(* IEC 61131-3 sources: moqui-plc/rust-plc/interfaces/codesys-iiot, 3 files *)

(* ---- json.st ---- *)
(* CODESYS IIoT JSON API used by moqui-plc (library namespace JSON).
 *
 * Interface declarations only (no implementation), for type checking with a
 * non-CODESYS compiler. The vendor library is object oriented (methods on
 * function blocks); the declarations mirror only the calls moqui-plc makes.
 *)

TYPE JSON_ERROR : (NO_ERROR, INVALID_INPUT, NO_MEMORY, NOT_FOUND, PARSE_ERROR); END_TYPE
TYPE JSONType : (JSON_OBJECT, JSON_ARRAY, KEY, VALUE); END_TYPE

TYPE JSONValue :
STRUCT
    wsValue : WSTRING(255);
    lrValue : LREAL;
    diValue : DINT;
    xValue : BOOL;
END_STRUCT
END_TYPE

TYPE JSONElement :
STRUCT
    eType : JSONType;
    diIndex : DINT;
    diParentIndex : DINT;
    value : JSONValue;
END_STRUCT
END_TYPE

FUNCTION_BLOCK JSONData
METHOD Clear
END_METHOD
METHOD GetElementByIndex : JSON_ERROR
VAR_INPUT
    diIndex : DINT;
END_VAR
VAR_OUTPUT
    jsonElement : JSONElement;
END_VAR
END_METHOD
METHOD GetChildren : JSON_ERROR
VAR_INPUT
    diIndex : DINT;
    pResult : POINTER TO JSONElement;
    udiMaxSize : UDINT;
END_VAR
VAR_OUTPUT
    udiResultSize : UDINT;
END_VAR
END_METHOD
END_FUNCTION_BLOCK

FUNCTION_BLOCK JSONDataFactory
METHOD Create : POINTER TO JSONData
VAR_OUTPUT
    eError : JSON_ERROR;
END_VAR
END_METHOD
END_FUNCTION_BLOCK

FUNCTION_BLOCK JSONBuilder
VAR_INPUT
    pJsonData : POINTER TO JSONData;
END_VAR
VAR_OUTPUT
    diRootObj : DINT;
END_VAR
METHOD Reset
END_METHOD
METHOD SetKeyWithObject : DINT
VAR_INPUT
    wsKey : WSTRING;
    diParentIndex : DINT;
END_VAR
END_METHOD
METHOD SetKeyWithValue : DINT
VAR_INPUT
    wsKey : WSTRING;
    value : ANY;
    diParentIndex : DINT;
END_VAR
END_METHOD
END_FUNCTION_BLOCK

FUNCTION_BLOCK JSONByteArrayWriter
VAR_INPUT
    xExecute : BOOL;
    xAsyncMode : BOOL;
    pwData : POINTER TO WORD;
    udiSize : UDINT;
    wsLineBreak : WSTRING(2);
END_VAR
VAR_IN_OUT
    jsonData : JSONData;
END_VAR
VAR_OUTPUT
    xDone : BOOL;
    xBusy : BOOL;
    xError : BOOL;
    eError : JSON_ERROR;
END_VAR
END_FUNCTION_BLOCK

FUNCTION_BLOCK JSONByteArrayReader
VAR_INPUT
    xExecute : BOOL;
    xAsyncMode : BOOL;
    pwData : POINTER TO WORD;
END_VAR
VAR_IN_OUT
    jsonData : JSONData;
END_VAR
VAR_OUTPUT
    xDone : BOOL;
    xBusy : BOOL;
    xError : BOOL;
    eError : JSON_ERROR;
END_VAR
END_FUNCTION_BLOCK

(* ---- mqtt.st ---- *)
(* CODESYS IIoT MQTT client API used by moqui-plc (library namespace MQTT).
 *
 * Interface declarations only (no implementation), for type checking with a
 * non-CODESYS compiler. Only the members moqui-plc uses are declared. A Rust
 * runtime would implement them on top of an MQTT 5 client crate.
 *)

TYPE MQTT_VERSION : (V3_1_1 := 4, V5 := 5); END_TYPE
TYPE MQTT_QOS : (QoS0, QoS1, QoS2); END_TYPE
TYPE MQTT_RETAIN_HANDLING : (On_Subscribe, If_Not_Exists, Not_Exists); END_TYPE
TYPE COMMUNICATION_MODE : (TCP, WEBSOCKET); END_TYPE
TYPE FILTER_MODE : (FILTER_OFF, FILTER_ON); END_TYPE
TYPE MQTT_ERROR : (NO_ERROR, TIMEOUT, CONNECTION_REFUSED, DISCONNECTED, PROTOCOL_ERROR); END_TYPE

(* Library parameters (CODESYS: MQTT.MQTTParam). Values are runtime specific. *)
VAR_GLOBAL CONSTANT
    g_udiMaxPacketSize : UDINT := 268435455;
    g_udiMaxUserProperties : UDINT := 8;
END_VAR

TYPE MQTTConnectProperties :
STRUCT
    udiSessionExpiryInterval : UDINT;
    udiMaximumPacketSize : UDINT;
END_STRUCT
END_TYPE

TYPE MQTTWillProperties :
STRUCT
    bPayloadFormatIndicator : BYTE;
    udiMessageExpiryInterval : UDINT;
    wsContentType : WSTRING;
    udiWillDelayInterval : UDINT;
END_STRUCT
END_TYPE

TYPE MQTTPublishProperties :
STRUCT
    bPayloadFormatIndicator : BYTE;
    udiMessageExpiryInterval : UDINT;
    wsContentType : WSTRING;
END_STRUCT
END_TYPE

TYPE MQTTSubscribeProperties :
STRUCT
    udiSubscriptionIdentifier : UDINT;
    xNoLocalOption : BOOL;
    xRetainAsPublished : BOOL;
    eRetainHandling : MQTT_RETAIN_HANDLING;
END_STRUCT
END_TYPE

FUNCTION_BLOCK MQTTClient
VAR_INPUT
    xEnable : BOOL;
    sHostname : STRING(255);
    uiPort : UINT;
    eCommunicationMode : COMMUNICATION_MODE;
    sWebSocketUrl : STRING(255);
    itfTLSContext : ITLSContext;
    eMQTTVersion : MQTT_VERSION;
    sClientId : STRING(255);
    wsUsername : WSTRING(255);
    wsPassword : WSTRING(255);
    uiKeepAlive : UINT;
    xCleanSession : BOOL;
    udiTimeOut : UDINT;
    tPingInterval : TIME;
    wsWillTopic : WSTRING(1024);
    pbWillMessage : POINTER TO BYTE;
    uiWillMessageSize : UINT;
    eWillQoS : MQTT_QOS;
    xWillRetain : BOOL;
    mQTTConnectProperties : MQTTConnectProperties;
    mQTTWillProperties : MQTTWillProperties;
END_VAR
VAR_OUTPUT
    xConnectedToBroker : BOOL;
    xBusy : BOOL;
    xError : BOOL;
    eMQTTError : MQTT_ERROR;
END_VAR
END_FUNCTION_BLOCK

FUNCTION_BLOCK MQTTPublish
VAR_INPUT
    xExecute : BOOL;
    mqttClient : REF_TO MQTTClient;
    wsTopicName : WSTRING(1024);
    pbPayload : POINTER TO BYTE;
    udiPayloadSize : UDINT;
    eQoS : MQTT_QOS;
    xRetain : BOOL;
    xReDelivery : BOOL;
    udiTimeOut : UDINT;
    mQTTPublishProperties : MQTTPublishProperties;
END_VAR
VAR_OUTPUT
    xDone : BOOL;
    xBusy : BOOL;
    xError : BOOL;
    eMQTTError : MQTT_ERROR;
END_VAR
END_FUNCTION_BLOCK

FUNCTION_BLOCK MQTTSubscribe
VAR_INPUT
    xEnable : BOOL;
    mqttClient : REF_TO MQTTClient;
    wsTopicFilter : WSTRING(1024);
    eFilterMode : FILTER_MODE;
    eSubscribeQoS : MQTT_QOS;
    pbPayload : POINTER TO BYTE;
    udiMaxPayloadSize : UDINT;
    udiTimeout : UDINT;
    mQTTSubscribeProperties : MQTTSubscribeProperties;
END_VAR
VAR_OUTPUT
    xDone : BOOL;
    xBusy : BOOL;
    xError : BOOL;
    eMQTTError : MQTT_ERROR;
    xSubscribeActive : BOOL;
    xReceived : BOOL;
    wsLastTopic : WSTRING(1024);
END_VAR
END_FUNCTION_BLOCK

(* ---- tls.st ---- *)
(* CODESYS Net Base Services TLS types used by moqui-plc (library namespace NBS).
 *
 * Interface declarations only (no implementation), for type checking with a
 * non-CODESYS compiler.
 *)

TYPE PURPOSE : (CLIENT_SIDE, SERVER_SIDE); END_TYPE

TYPE CIPHER_LIST :
STRUCT
    psList : POINTER TO STRING;
    udiSize : UDINT;
END_STRUCT
END_TYPE

TYPE CERT_INFO :
STRUCT
    psInfo : POINTER TO STRING;
    udiSize : UDINT;
END_STRUCT
END_TYPE

(* CODESYS passes the TLS context as an interface; 0 means no TLS. *)
TYPE ITLSContext : POINTER TO TLSContext; END_TYPE

FUNCTION_BLOCK TLSContext
VAR_INPUT
    sUseCaseName : STRING;
    ePurpose : PURPOSE;
    sTLSVersion : STRING;
    sCipherList : CIPHER_LIST;
    sHostname : STRING(255);
    ciCertInfo : CERT_INFO;
    udiVerificationMode : UDINT;
    itfCertVerifer : LWORD; (* certificate verifier interface; 0 = none *)
END_VAR
END_FUNCTION_BLOCK
